// SIMATIC S7-200 project (STEP 7-Micro/WIN), CPU 224 CN REL 02.01

SYMBOL_TABLE USUARIO1
SB1R             I1.3     // Pulsador de marcha (verde)
SB2R             I1.2     // Pulsador de paro (rojo)
SA               I1.5     // Selector de modo
QSR              I1.4     // Zeta de emergencia
SM1R             I0.3     // Cilindro largo retraido
SM2R             I0.2     // Cilindro largo extendido
SM3R             I0.1     // Pinza de dedo cerrado
SM4R             I0.4     // Cilindro delgado retraido
SM5R             I0.5     // Cilindro delgado extendido
SF1R             I0.0     // Sensor optico
KB1R             Q0.2     // Accionamiento del cilindro largo
KB2R             Q0.0     // Accionamiento de la pinza
KB3R             Q0.3     // Accionamiento del cilindro delgado
HL1R             Q0.7     // Piloto indicador  de parada
HL2R             Q1.0     // Piloto indicador de marcha
HL3R             Q1.1     // Piloto indicador de emergencia
E0               M0.0     // Estado inicial
E1               M0.1     // Estado para el cierre de la pinza neumatica
E2               M0.2     // Estado para el retroceso del cilindro largo
E3               M0.3     // Estado de salida del cilindro delgado
E4               M0.4     // Estado de retroceso del cilindro delgado
E5               M0.5     // Estado de extension del cilindro largo
E6               M0.6     // Estado de apertura de la garra y avisos
EM               M1.0     // Estado de emergencia
EM1              M1.1     // Estado para la apertura de la garra
EM2              M1.2     // Estado auxiliar para el retorno al estado inicial
EP               M1.3     // Estado de parada
END_SYMBOL_TABLE

ORGANIZATION_BLOCK PRINCIPAL:OB1
TITLE=COMENTARIOS DEL PROGRAMA
BEGIN
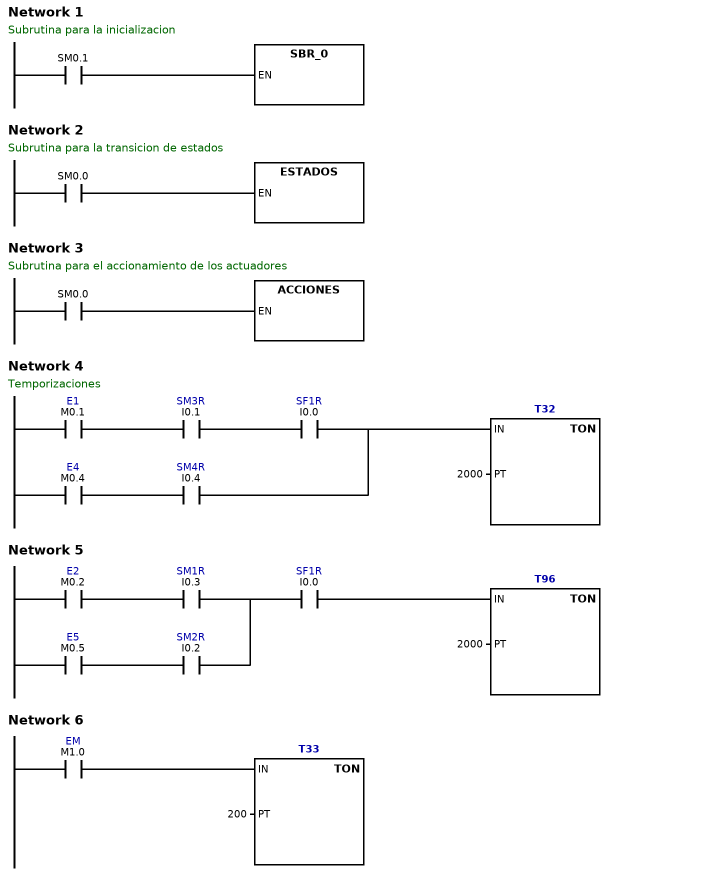
Network 1
// Subrutina para la inicializacion
LD     SM0.1
CALL   SBR_0:SBR0
Network 2
// Subrutina para la transicion de estados
LD     SM0.0
CALL   ESTADOS:SBR1
Network 3
// Subrutina para el accionamiento de los actuadores
LD     SM0.0
CALL   ACCIONES:SBR2
Network 4
// Temporizaciones
LD     E1:M0.1
A      SM3R:I0.1
A      SF1R:I0.0
LD     E4:M0.4
A      SM4R:I0.4
OLD
TON    T32, 2000
Network 5
LD     E2:M0.2
A      SM1R:I0.3
LD     E5:M0.5
A      SM2R:I0.2
OLD
A      SF1R:I0.0
TON    T96, 2000
Network 6
LD     EM:M1.0
TON    T33, 200
END_ORGANIZATION_BLOCK

SUBROUTINE_BLOCK SBR_0:SBR0
TITLE=COMENTARIOS DE LA SUBRUTINA
BEGIN
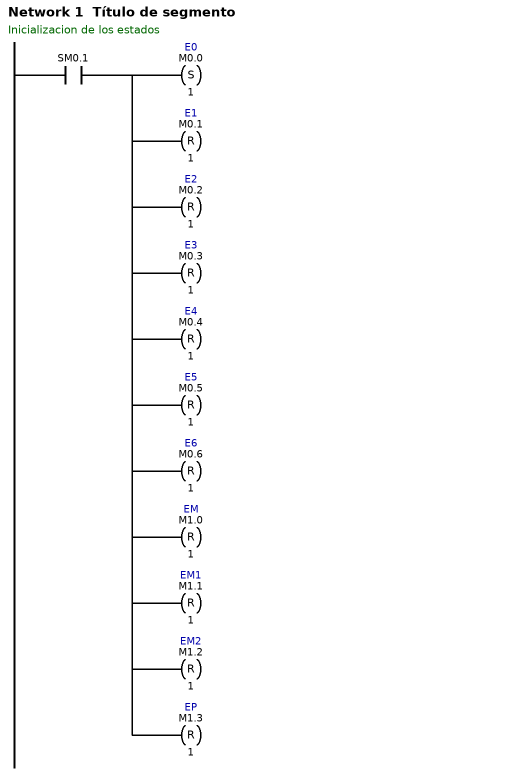
Network 1 // Título de segmento
// Inicializacion de los estados
LD     SM0.1
S      E0:M0.0, 1
R      E1:M0.1, 1
R      E2:M0.2, 1
R      E3:M0.3, 1
R      E4:M0.4, 1
R      E5:M0.5, 1
R      E6:M0.6, 1
R      EM:M1.0, 1
R      EM1:M1.1, 1
R      EM2:M1.2, 1
R      EP:M1.3, 1
END_SUBROUTINE_BLOCK

SUBROUTINE_BLOCK ESTADOS:SBR1
TITLE=TRANSICION DE ESTADOS
BEGIN
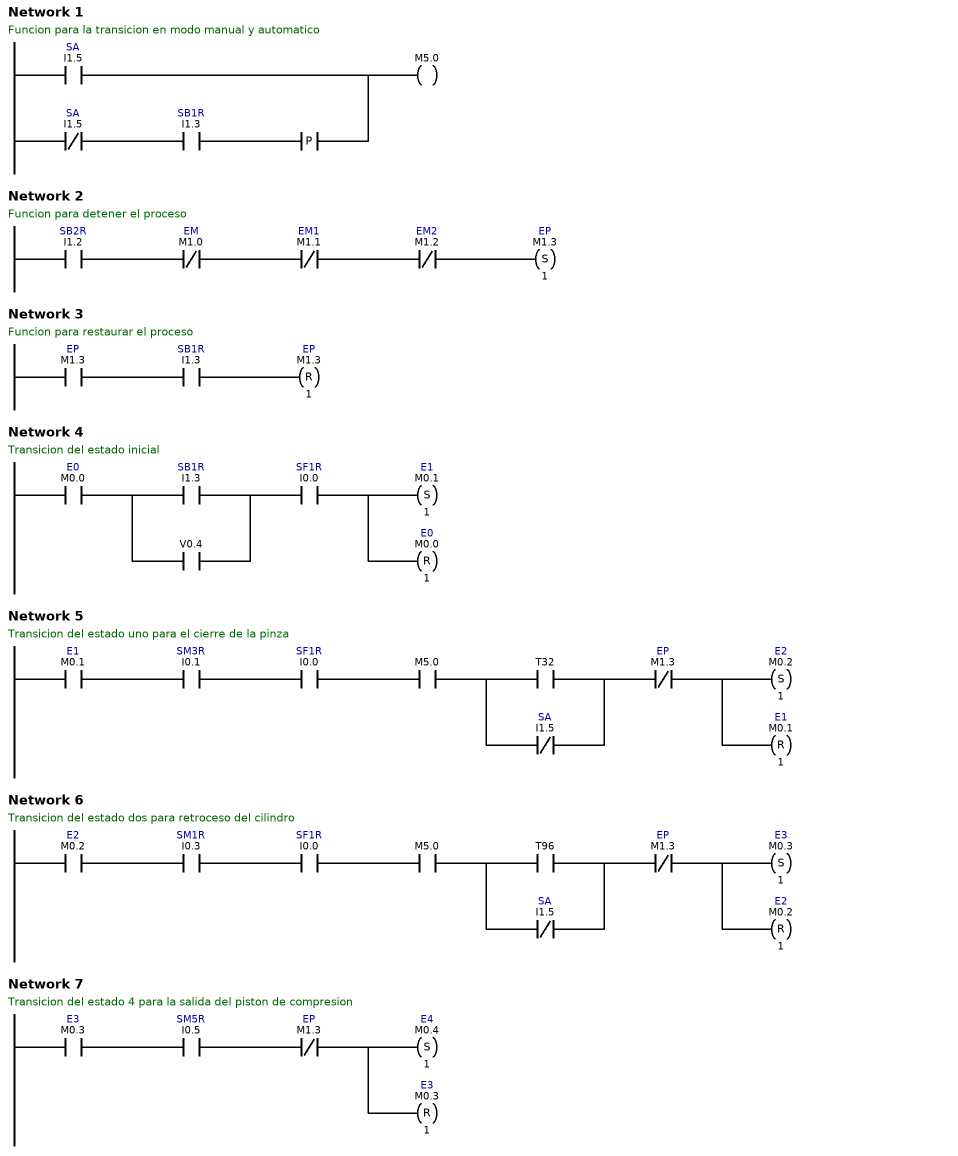
Network 1
// Funcion para la transicion en modo manual y automatico
LD     SA:I1.5
LDN    SA:I1.5
A      SB1R:I1.3
EU
OLD
=      M5.0
Network 2
// Funcion para detener el proceso
LD     SB2R:I1.2
AN     EM:M1.0
AN     EM1:M1.1
AN     EM2:M1.2
S      EP:M1.3, 1
Network 3
// Funcion para restaurar el proceso
LD     EP:M1.3
A      SB1R:I1.3
R      EP:M1.3, 1
Network 4
// Transicion del estado inicial
LD     E0:M0.0
LD     SB1R:I1.3
O      V0.4
ALD
A      SF1R:I0.0
S      E1:M0.1, 1
R      E0:M0.0, 1
Network 5
// Transicion del estado uno para el cierre de la pinza
LD     E1:M0.1
A      SM3R:I0.1
A      SF1R:I0.0
A      M5.0
LD     T32
ON     SA:I1.5
ALD
AN     EP:M1.3
S      E2:M0.2, 1
R      E1:M0.1, 1
Network 6
// Transicion del estado dos para retroceso del cilindro
LD     E2:M0.2
A      SM1R:I0.3
A      SF1R:I0.0
A      M5.0
LD     T96
ON     SA:I1.5
ALD
AN     EP:M1.3
S      E3:M0.3, 1
R      E2:M0.2, 1
Network 7
// Transicion del estado 4 para la salida del piston de compresion
LD     E3:M0.3
A      SM5R:I0.5
AN     EP:M1.3
S      E4:M0.4, 1
R      E3:M0.3, 1
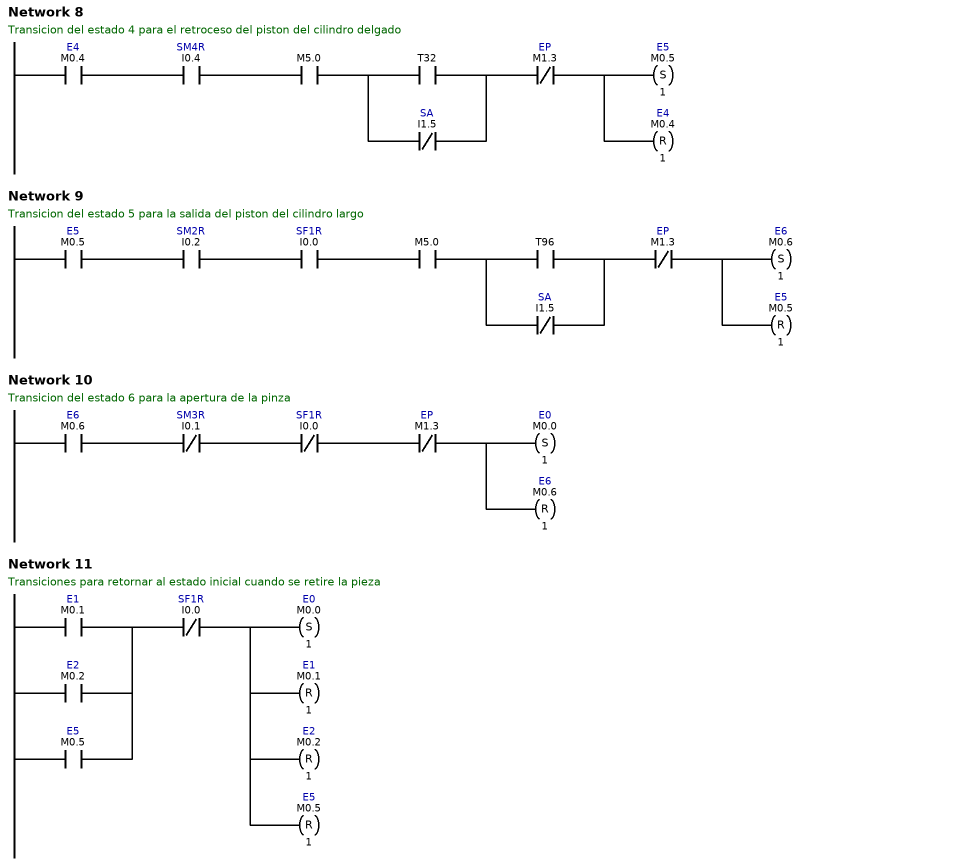
Network 8
// Transicion del estado 4 para el retroceso del piston del cilindro delgado
LD     E4:M0.4
A      SM4R:I0.4
A      M5.0
LD     T32
ON     SA:I1.5
ALD
AN     EP:M1.3
S      E5:M0.5, 1
R      E4:M0.4, 1
Network 9
// Transicion del estado 5 para la salida del piston del cilindro largo
LD     E5:M0.5
A      SM2R:I0.2
A      SF1R:I0.0
A      M5.0
LD     T96
ON     SA:I1.5
ALD
AN     EP:M1.3
S      E6:M0.6, 1
R      E5:M0.5, 1
Network 10
// Transicion del estado 6 para la apertura de la pinza
LD     E6:M0.6
AN     SM3R:I0.1
AN     SF1R:I0.0
AN     EP:M1.3
S      E0:M0.0, 1
R      E6:M0.6, 1
Network 11
// Transiciones para retornar al estado inicial cuando se retire la pieza
LD     E1:M0.1
O      E2:M0.2
O      E5:M0.5
AN     SF1R:I0.0
S      E0:M0.0, 1
R      E1:M0.1, 1
R      E2:M0.2, 1
R      E5:M0.5, 1
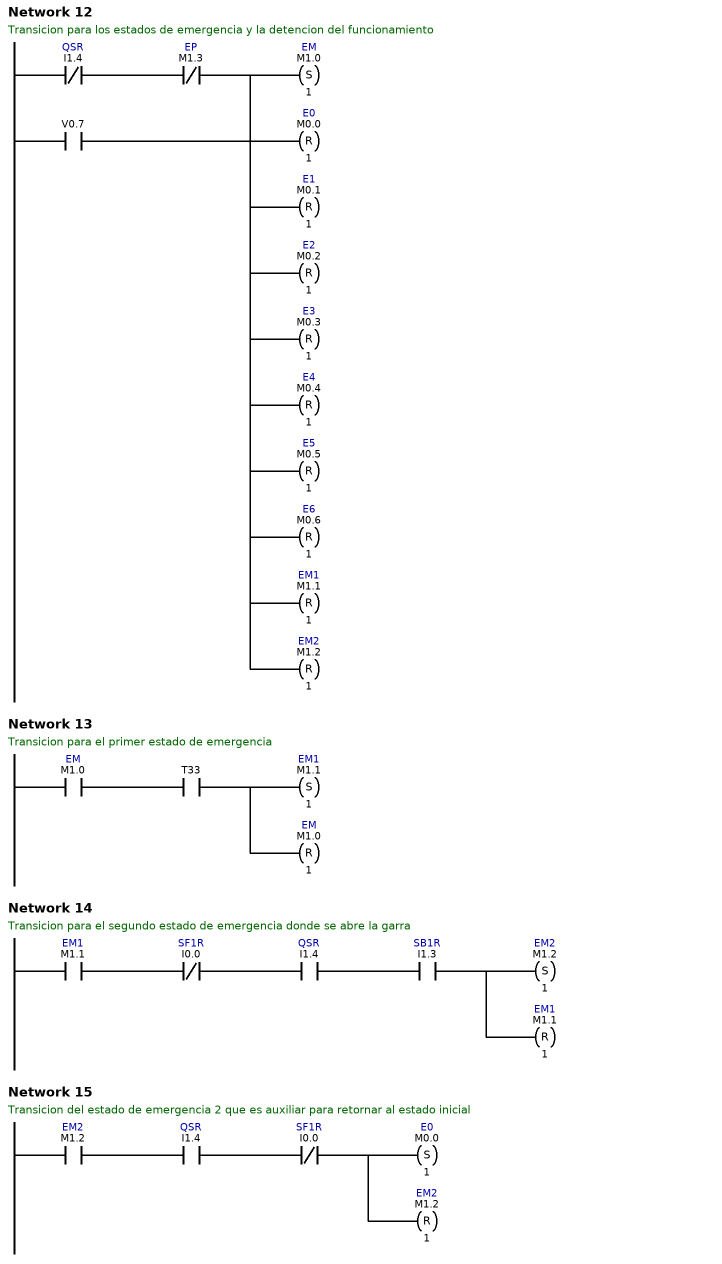
Network 12
// Transicion para los estados de emergencia y la detencion del funcionamiento
LDN    QSR:I1.4
AN     EP:M1.3
O      V0.7
S      EM:M1.0, 1
R      E0:M0.0, 1
R      E1:M0.1, 1
R      E2:M0.2, 1
R      E3:M0.3, 1
R      E4:M0.4, 1
R      E5:M0.5, 1
R      E6:M0.6, 1
R      EM1:M1.1, 1
R      EM2:M1.2, 1
Network 13
// Transicion para el primer estado de emergencia
LD     EM:M1.0
A      T33
S      EM1:M1.1, 1
R      EM:M1.0, 1
Network 14
// Transicion para el segundo estado de emergencia donde se abre la garra
LD     EM1:M1.1
AN     SF1R:I0.0
A      QSR:I1.4
A      SB1R:I1.3
S      EM2:M1.2, 1
R      EM1:M1.1, 1
Network 15
// Transicion del estado de emergencia 2 que es auxiliar para retornar al estado inicial
LD     EM2:M1.2
A      QSR:I1.4
AN     SF1R:I0.0
S      E0:M0.0, 1
R      EM2:M1.2, 1
END_SUBROUTINE_BLOCK

SUBROUTINE_BLOCK ACCIONES:SBR2
TITLE=SUBRUTINA PARA EL ACCIONAMIENTO DE LOS ACTUADORES
BEGIN
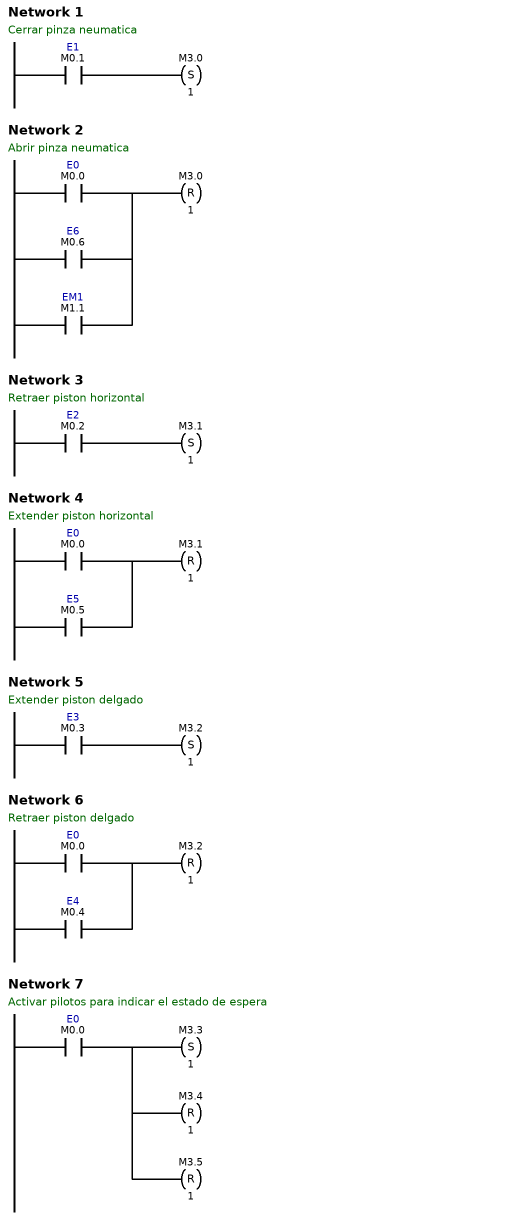
Network 1
// Cerrar pinza neumatica
LD     E1:M0.1
S      M3.0, 1
Network 2
// Abrir pinza neumatica
LD     E0:M0.0
O      E6:M0.6
O      EM1:M1.1
R      M3.0, 1
Network 3
// Retraer piston horizontal
LD     E2:M0.2
S      M3.1, 1
Network 4
// Extender piston horizontal
LD     E0:M0.0
O      E5:M0.5
R      M3.1, 1
Network 5
// Extender piston delgado
LD     E3:M0.3
S      M3.2, 1
Network 6
// Retraer piston delgado
LD     E0:M0.0
O      E4:M0.4
R      M3.2, 1
Network 7
// Activar pilotos para indicar el estado de espera
LD     E0:M0.0
S      M3.3, 1
R      M3.4, 1
R      M3.5, 1
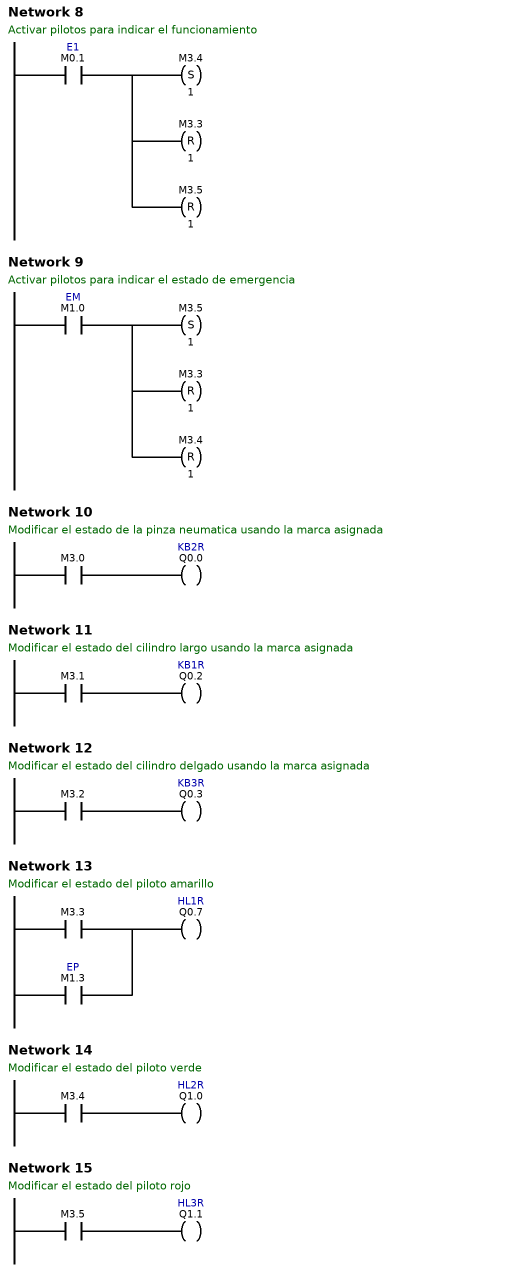
Network 8
// Activar pilotos para indicar el funcionamiento
LD     E1:M0.1
S      M3.4, 1
R      M3.3, 1
R      M3.5, 1
Network 9
// Activar pilotos para indicar el estado de emergencia
LD     EM:M1.0
S      M3.5, 1
R      M3.3, 1
R      M3.4, 1
Network 10
// Modificar el estado de la pinza neumatica usando la marca asignada
LD     M3.0
=      KB2R:Q0.0
Network 11
// Modificar el estado del cilindro largo usando la marca asignada
LD     M3.1
=      KB1R:Q0.2
Network 12
// Modificar el estado del cilindro delgado usando la marca asignada
LD     M3.2
=      KB3R:Q0.3
Network 13
// Modificar el estado del piloto amarillo
LD     M3.3
O      EP:M1.3
=      HL1R:Q0.7
Network 14
// Modificar el estado del piloto verde
LD     M3.4
=      HL2R:Q1.0
Network 15
// Modificar el estado del piloto rojo
LD     M3.5
=      HL3R:Q1.1
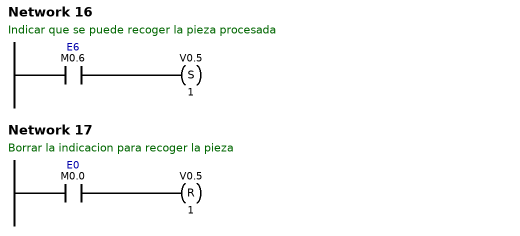
Network 16
// Indicar que se puede recoger la pieza procesada
LD     E6:M0.6
S      V0.5, 1
Network 17
// Borrar la indicacion para recoger la pieza 
LD     E0:M0.0
R      V0.5, 1
END_SUBROUTINE_BLOCK
